ABB RAPID module: Long_ProgramName12.mod

MODULE MOD_Long_ProgramName12

PERS wobjdata rdkWObj := [FALSE, TRUE, "", [[0,0,0],[1,0,0,0]],[[0,0,0],[1,0,0,0]]];
PERS tooldata rdkTool := [TRUE,[[0,0,0],[1,0,0,0]],[6.8,[0,0,15],[1,0,0,0],0,0,0.005]];
VAR speeddata rdkSpeed := [500,500,500,500];
VAR zonedata rdkZone := z1;
VAR extjoint rdkExtax := [9E9,9E9,9E9,9E9,9E9,9E9];

PROC main_RoboDK()
	Long_ProgramName12;
	EXIT;
ENDPROC

PROC Long_ProgramName12()
	!Program generated by RoboDK v5.9.4 for ABB IRB 1600-8/1.45 on 26/10/2026 01:01:07
	!Using nominal kinematics.
	var robtarget crt;
	crt := CRobT(\Tool:=rdkTool, \WObj:=rdkWObj);
	rdkExtax := crt.extax;
	ConfJ \On;
	ConfL \Off;
	!Long body
	rdkTool.tframe:=[[10.000,0.000,150.000],[1.00000000,0.00000000,0.00000000,0.00000000]];
	MoveL [[40.000,40.000,0.000],[0.58801837,0.20533497,0.76632048,-0.15755906],[-1,-1,0,1],rdkExtax], rdkSpeed, rdkZone, rdkTool, \WObj:=rdkWObj;
ENDPROC

ENDMODULE
